Fanuc KAREL source: KO00023.KL

PROGRAM KO00023
%NOLOCKGROUP
VAR
  P1: XYZWPREXT
  P2: XYZWPREXT
  P3: XYZWPREXT
  P4: XYZWPREXT
  OUT: XYZWPREXT
BEGIN
  OUT = FRAME(P1, P2, P3, P4)
END KO00023
